Fanuc KAREL source: kd00008.KL

PROGRAM KD00008
%STACKSIZE=65535
%PRIORITY=65535
%TPMOTION
%NOLOCKGROUP
VAR
I : INTEGER
J : INTEGER
B : BOOLEAN
R : REAL
S : STRING[80]
BEGIN
I=1
END KD00008
